// Mitsubishi GX Works2 project: 261019_적산 타이머 실습_타이머 추가 응용1   PLC: Q03UDV

PROGRAM MAIN
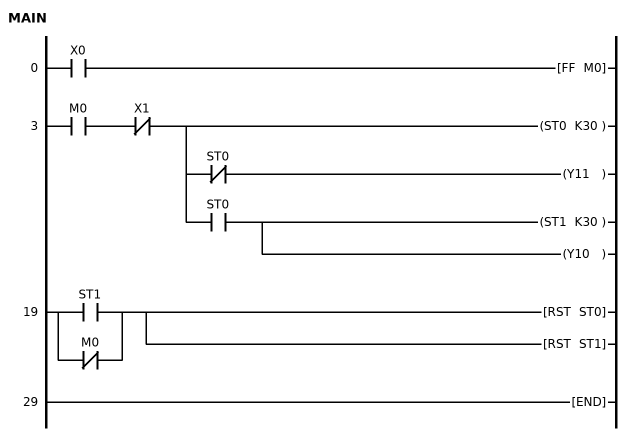
0     LD      X0
      FF      M0
3     LD      M0
      ANI     X1
      OUT     ST0 K30
      MPS
      ANI     ST0
      OUT     Y11
      MPP
      AND     ST0
      OUT     ST1 K30
      OUT     Y10
19    LD      ST1
      ORI     M0
      RST     ST0
      RST     ST1
29    END
END_PROGRAM
